// TIA Portal V20 export
// export: Created 2026-10-19T18:36:00.5112629Z, ExportSetting WithDefaults, DisplayName Totally Integrated Automation Portal, DisplayVersion V20 Update 6, DisplayName TIA Portal Openness, DisplayVersion V20 Update 6, DisplayName TIA Portal Version Control Interface, DisplayVersion V20 Update 6, DisplayName SINAMICS Startdrive Advanced, DisplayVersion V20 SP1, DisplayName SINAMICS Startdrive G130, G150, S120, S150, SINAMICS MV, G220, S200, S210, DisplayVersion V20 SP1, DisplayName SINAMICS Startdrive G110M, G120, G120C, G120D, G120P, G115D, DisplayVersion V20 SP1, DisplayName STEP 7 Professional, DisplayVersion V20 Update 6, DisplayName STEP 7 Safety, DisplayVersion V20 Update 2, DisplayName WinCC Basic/Comfort/Advanced, DisplayVersion V20 Update 6, DisplayName WinCC Unified, DisplayVersion V20 Update 6
FUNCTION_BLOCK "Main_Safety_RTG1"   // FB1, F_FBD
{ S7_Optimized_Access := 'TRUE' }
VERSION : 0.1
// stored: AutoNumber false, IsIECCheckEnabled false, UDAEnableTagReadback false
   VAR
      Safety_OK : Bool;
   END_VAR
   VAR_TEMP
      HMI_1_Estop_Pressed_1 : Bool;
      HMI_1_Estop_Pressed_2 : Bool;
      HMI_2_Estop_Pressed_1 : Bool;
      HMI_2_Estop_Pressed_2 : Bool;
      HMI_1_Reset_Comiss_1 : Bool;
      HMI_1_Reset_Comiss_2 : Bool;
      HMI_2_Reset_Comiss_1 : Bool;
      HMI_2_Reset_Comiss_2 : Bool;
   END_VAR
BEGIN

REGION Network 1: HMI 1 EMERGENCY BUTTON AND RESET COMISSIONING
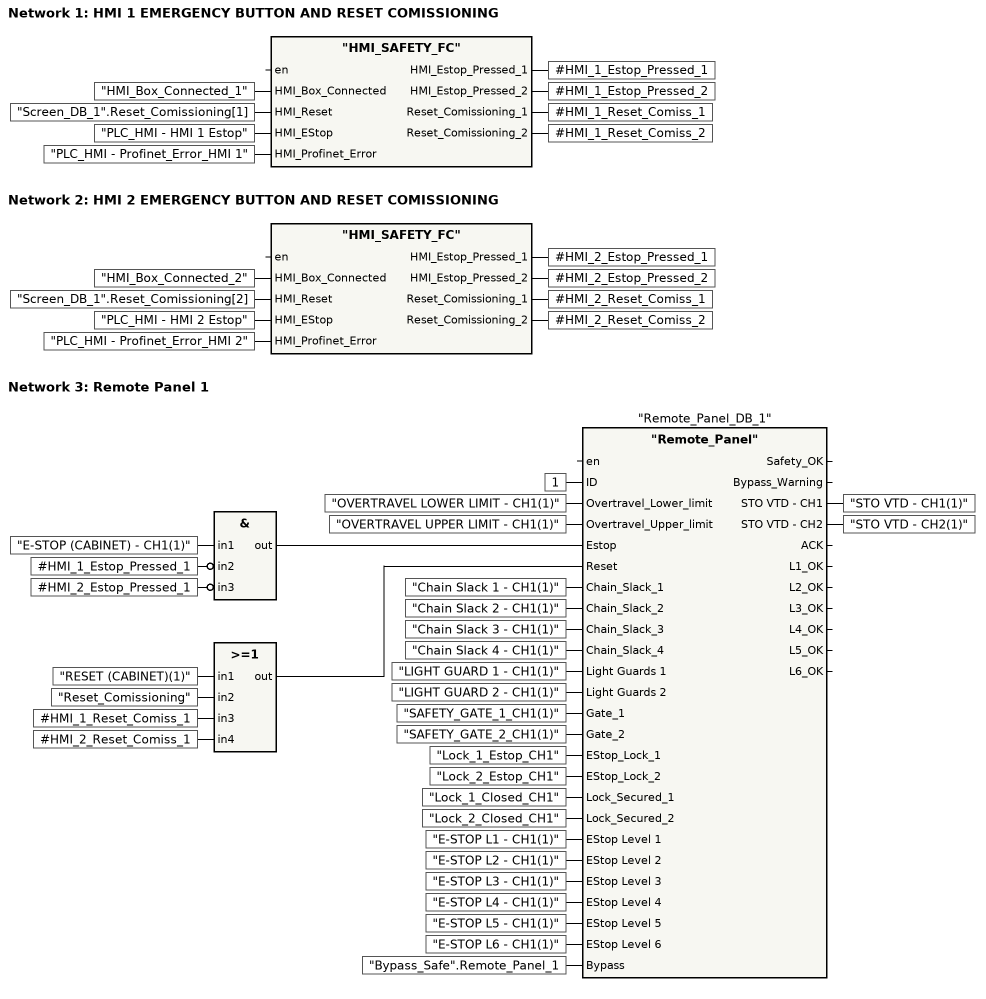
   "HMI_SAFETY_FC"(HMI_Box_Connected := "HMI_Box_Connected_1",
                   HMI_Reset := "Screen_DB_1".Reset_Comissioning[1],
                   HMI_EStop := "PLC_HMI - HMI 1 Estop",
                   HMI_Profinet_Error := "PLC_HMI - Profinet_Error_HMI 1",
                   HMI_Estop_Pressed_1 => #HMI_1_Estop_Pressed_1,
                   HMI_Estop_Pressed_2 => #HMI_1_Estop_Pressed_2,
                   Reset_Comissioning_1 => #HMI_1_Reset_Comiss_1,
                   Reset_Comissioning_2 => #HMI_1_Reset_Comiss_2);
END_REGION

REGION Network 2: HMI 2 EMERGENCY BUTTON AND RESET COMISSIONING
   "HMI_SAFETY_FC"(HMI_Box_Connected := "HMI_Box_Connected_2",
                   HMI_Reset := "Screen_DB_1".Reset_Comissioning[2],
                   HMI_EStop := "PLC_HMI - HMI 2 Estop",
                   HMI_Profinet_Error := "PLC_HMI - Profinet_Error_HMI 2",
                   HMI_Estop_Pressed_1 => #HMI_2_Estop_Pressed_1,
                   HMI_Estop_Pressed_2 => #HMI_2_Estop_Pressed_2,
                   Reset_Comissioning_1 => #HMI_2_Reset_Comiss_1,
                   Reset_Comissioning_2 => #HMI_2_Reset_Comiss_2);
END_REGION

REGION Network 3: Remote Panel 1
   "Remote_Panel_DB_1"(ID := 1,   // "Remote_Panel"
                       Overtravel_Lower_limit := "OVERTRAVEL LOWER LIMIT - CH1(1)",
                       Overtravel_Upper_limit := "OVERTRAVEL UPPER LIMIT - CH1(1)",
                       Estop := "E-STOP (CABINET) - CH1(1)" AND NOT #HMI_1_Estop_Pressed_1 AND NOT #HMI_2_Estop_Pressed_1,
                       Reset := "RESET (CABINET)(1)" OR "Reset_Comissioning" OR #HMI_1_Reset_Comiss_1 OR #HMI_2_Reset_Comiss_1,
                       Chain_Slack_1 := "Chain Slack 1 - CH1(1)",
                       Chain_Slack_2 := "Chain Slack 2 - CH1(1)",
                       Chain_Slack_3 := "Chain Slack 3 - CH1(1)",
                       Chain_Slack_4 := "Chain Slack 4 - CH1(1)",
                       "Light Guards 1" := "LIGHT GUARD 1 - CH1(1)",
                       "Light Guards 2" := "LIGHT GUARD 2 - CH1(1)",
                       Gate_1 := "SAFETY_GATE_1_CH1(1)",
                       Gate_2 := "SAFETY_GATE_2_CH1(1)",
                       EStop_Lock_1 := "Lock_1_Estop_CH1",
                       EStop_Lock_2 := "Lock_2_Estop_CH1",
                       Lock_Secured_1 := "Lock_1_Closed_CH1",
                       Lock_Secured_2 := "Lock_2_Closed_CH1",
                       "EStop Level 1" := "E-STOP L1 - CH1(1)",
                       "EStop Level 2" := "E-STOP L2 - CH1(1)",
                       "EStop Level 3" := "E-STOP L3 - CH1(1)",
                       "EStop Level 4" := "E-STOP L4 - CH1(1)",
                       "EStop Level 5" := "E-STOP L5 - CH1(1)",
                       "EStop Level 6" := "E-STOP L6 - CH1(1)",
                       Bypass := "Bypass_Safe".Remote_Panel_1,
                       "STO VTD - CH1" => "STO VTD - CH1(1)",
                       "STO VTD - CH2" => "STO VTD - CH2(1)");
END_REGION

REGION Network 4: Remote Panel 2
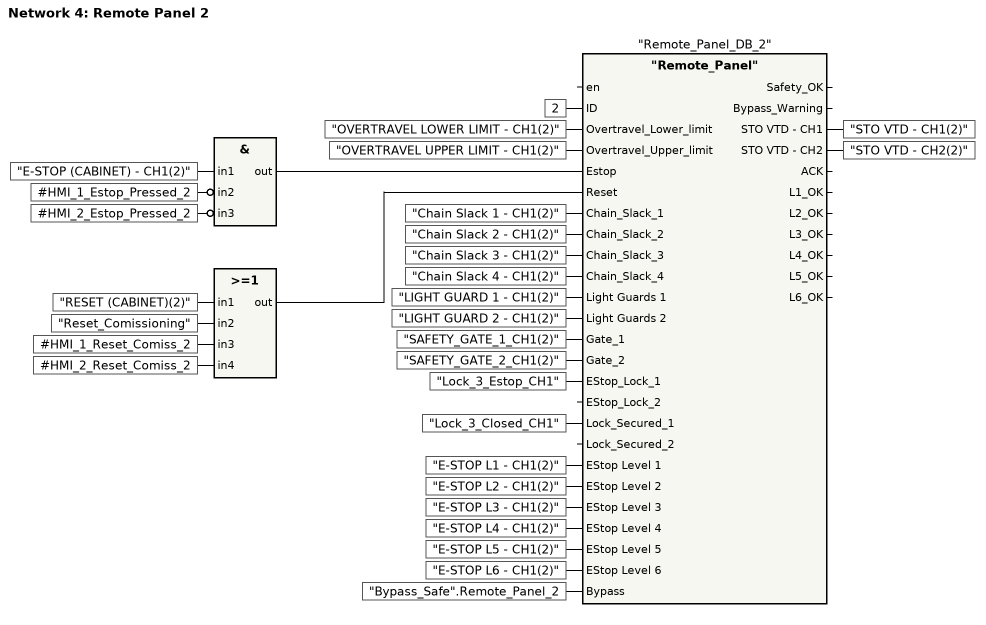
   "Remote_Panel_DB_2"(ID := 2,   // "Remote_Panel"
                       Overtravel_Lower_limit := "OVERTRAVEL LOWER LIMIT - CH1(2)",
                       Overtravel_Upper_limit := "OVERTRAVEL UPPER LIMIT - CH1(2)",
                       Estop := "E-STOP (CABINET) - CH1(2)" AND NOT #HMI_1_Estop_Pressed_2 AND NOT #HMI_2_Estop_Pressed_2,
                       Reset := "RESET (CABINET)(2)" OR "Reset_Comissioning" OR #HMI_1_Reset_Comiss_2 OR #HMI_2_Reset_Comiss_2,
                       Chain_Slack_1 := "Chain Slack 1 - CH1(2)",
                       Chain_Slack_2 := "Chain Slack 2 - CH1(2)",
                       Chain_Slack_3 := "Chain Slack 3 - CH1(2)",
                       Chain_Slack_4 := "Chain Slack 4 - CH1(2)",
                       "Light Guards 1" := "LIGHT GUARD 1 - CH1(2)",
                       "Light Guards 2" := "LIGHT GUARD 2 - CH1(2)",
                       Gate_1 := "SAFETY_GATE_1_CH1(2)",
                       Gate_2 := "SAFETY_GATE_2_CH1(2)",
                       EStop_Lock_1 := "Lock_3_Estop_CH1",
                       Lock_Secured_1 := "Lock_3_Closed_CH1",
                       "EStop Level 1" := "E-STOP L1 - CH1(2)",
                       "EStop Level 2" := "E-STOP L2 - CH1(2)",
                       "EStop Level 3" := "E-STOP L3 - CH1(2)",
                       "EStop Level 4" := "E-STOP L4 - CH1(2)",
                       "EStop Level 5" := "E-STOP L5 - CH1(2)",
                       "EStop Level 6" := "E-STOP L6 - CH1(2)",
                       Bypass := "Bypass_Safe".Remote_Panel_2,
                       "STO VTD - CH1" => "STO VTD - CH1(2)",
                       "STO VTD - CH2" => "STO VTD - CH2(2)");
END_REGION

REGION Network 5: ESTOP LEVEL PANELS
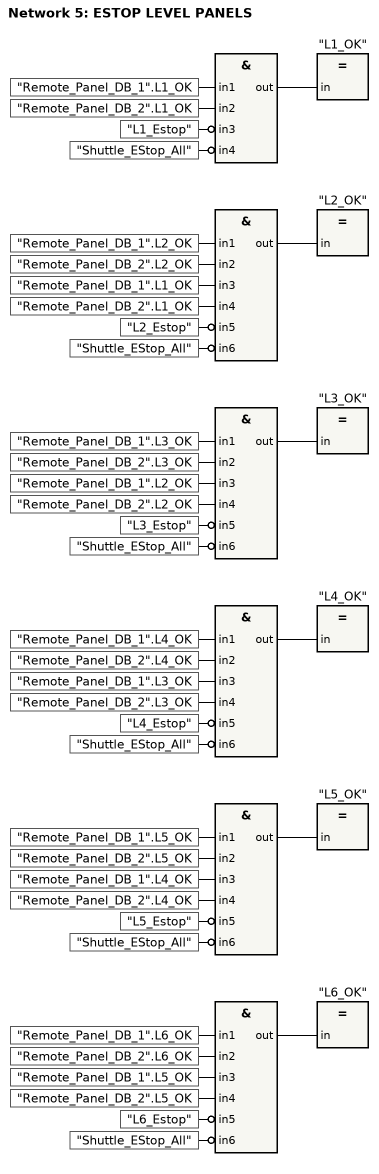
   "L1_OK" := "Remote_Panel_DB_1".L1_OK AND "Remote_Panel_DB_2".L1_OK AND NOT "L1_Estop" AND NOT "Shuttle_EStop_All";
   "L2_OK" := "Remote_Panel_DB_1".L2_OK AND "Remote_Panel_DB_2".L2_OK AND "Remote_Panel_DB_1".L1_OK AND "Remote_Panel_DB_2".L1_OK AND NOT "L2_Estop" AND NOT "Shuttle_EStop_All";
   "L3_OK" := "Remote_Panel_DB_1".L3_OK AND "Remote_Panel_DB_2".L3_OK AND "Remote_Panel_DB_1".L2_OK AND "Remote_Panel_DB_2".L2_OK AND NOT "L3_Estop" AND NOT "Shuttle_EStop_All";
   "L4_OK" := "Remote_Panel_DB_1".L4_OK AND "Remote_Panel_DB_2".L4_OK AND "Remote_Panel_DB_1".L3_OK AND "Remote_Panel_DB_2".L3_OK AND NOT "L4_Estop" AND NOT "Shuttle_EStop_All";
   "L5_OK" := "Remote_Panel_DB_1".L5_OK AND "Remote_Panel_DB_2".L5_OK AND "Remote_Panel_DB_1".L4_OK AND "Remote_Panel_DB_2".L4_OK AND NOT "L5_Estop" AND NOT "Shuttle_EStop_All";
   "L6_OK" := "Remote_Panel_DB_1".L6_OK AND "Remote_Panel_DB_2".L6_OK AND "Remote_Panel_DB_1".L5_OK AND "Remote_Panel_DB_2".L5_OK AND NOT "L6_Estop" AND NOT "Shuttle_EStop_All";
END_REGION

REGION Network 6: LOCKS
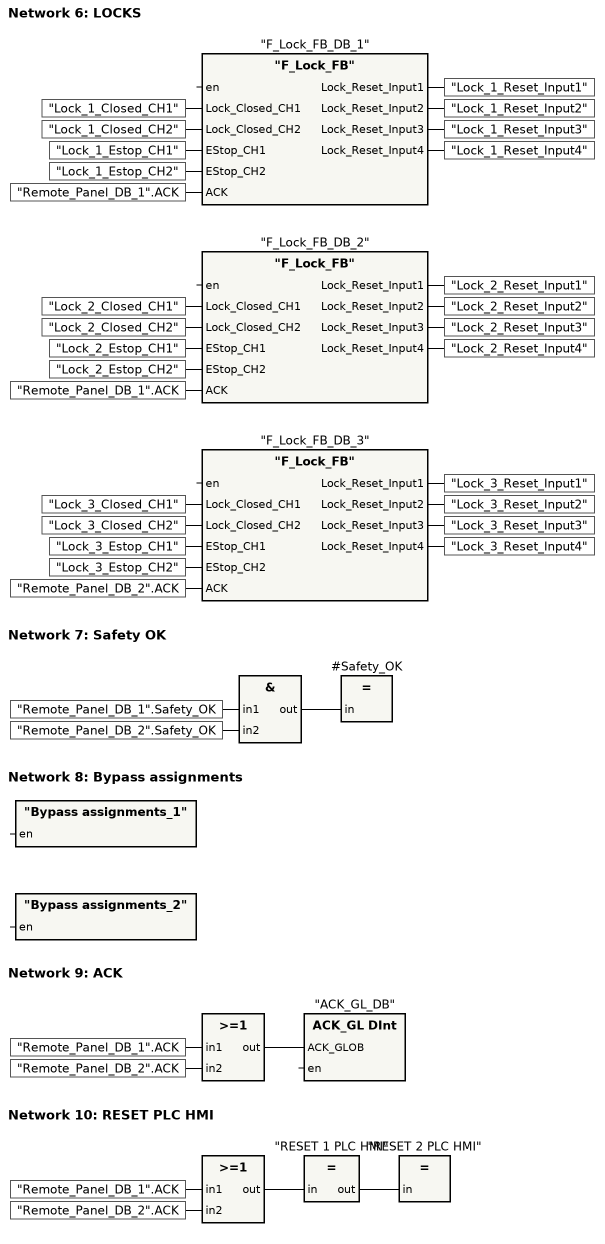
   "F_Lock_FB_DB_1"(Lock_Closed_CH1 := "Lock_1_Closed_CH1",   // "F_Lock_FB"
                    Lock_Closed_CH2 := "Lock_1_Closed_CH2",
                    EStop_CH1 := "Lock_1_Estop_CH1",
                    EStop_CH2 := "Lock_1_Estop_CH2",
                    ACK := "Remote_Panel_DB_1".ACK,
                    Lock_Reset_Input1 => "Lock_1_Reset_Input1",
                    Lock_Reset_Input2 => "Lock_1_Reset_Input2",
                    Lock_Reset_Input3 => "Lock_1_Reset_Input3",
                    Lock_Reset_Input4 => "Lock_1_Reset_Input4");
   "F_Lock_FB_DB_2"(Lock_Closed_CH1 := "Lock_2_Closed_CH1",   // "F_Lock_FB"
                    Lock_Closed_CH2 := "Lock_2_Closed_CH2",
                    EStop_CH1 := "Lock_2_Estop_CH1",
                    EStop_CH2 := "Lock_2_Estop_CH2",
                    ACK := "Remote_Panel_DB_1".ACK,
                    Lock_Reset_Input1 => "Lock_2_Reset_Input1",
                    Lock_Reset_Input2 => "Lock_2_Reset_Input2",
                    Lock_Reset_Input3 => "Lock_2_Reset_Input3",
                    Lock_Reset_Input4 => "Lock_2_Reset_Input4");
   "F_Lock_FB_DB_3"(Lock_Closed_CH1 := "Lock_3_Closed_CH1",   // "F_Lock_FB"
                    Lock_Closed_CH2 := "Lock_3_Closed_CH2",
                    EStop_CH1 := "Lock_3_Estop_CH1",
                    EStop_CH2 := "Lock_3_Estop_CH2",
                    ACK := "Remote_Panel_DB_2".ACK,
                    Lock_Reset_Input1 => "Lock_3_Reset_Input1",
                    Lock_Reset_Input2 => "Lock_3_Reset_Input2",
                    Lock_Reset_Input3 => "Lock_3_Reset_Input3",
                    Lock_Reset_Input4 => "Lock_3_Reset_Input4");
END_REGION

REGION Network 7: Safety OK
   #Safety_OK := "Remote_Panel_DB_1".Safety_OK AND "Remote_Panel_DB_2".Safety_OK;
END_REGION

REGION Network 8: Bypass assignments
   "Bypass assignments_1"();
   "Bypass assignments_2"();
END_REGION

REGION Network 9: ACK
   "ACK_GL_DB"(ACK_GLOB := "Remote_Panel_DB_1".ACK OR "Remote_Panel_DB_2".ACK);   // ACK_GL
END_REGION

REGION Network 10: RESET PLC HMI
   "RESET 1 PLC HMI" := "Remote_Panel_DB_1".ACK OR "Remote_Panel_DB_2".ACK;
   "RESET 2 PLC HMI" := "RESET 1 PLC HMI";
END_REGION
END_FUNCTION_BLOCK
